(* IEC 61131-3 sources: 2026_Projet_YGO_ExcavatriceDragage/CODE_BACKUP/CODE_20260904_AvantWeekendBackup_v0.6.34/H_TREUILS_BENNE/_TYPES, 19 files *)

(* ---- E_WinchFinalInterlockReason.st ---- *)
(* =======================================================================
   🔒 E_WinchFinalInterlockReason — Raisons de blocage barrière finale
   ───────────────────────────────────────────────────────────────
   🎯 Rôle : Énumération des causes de neutralisation/interlock final treuil
   📄 Doc métier : DOC/AF/AF_Partie-10_Fonction_Winch_v2.1.md
   ======================================================================= *)
{attribute 'qualified_only'}
TYPE E_WinchFinalInterlockReason :
(
    NONE                        := 0,                                 // Aucun blocage actif
    BRAKE_COMMAND_NOT_CONFIRMED := 1,                                 // Absence confirmation ouverture frein > 500ms
    RESTART_INHIBITED           := 2,                                 // Inhibition redemarrage actif
    SENSE_DROP_TIMEOUT          := 3                                  // T_max §3bis depasse sans confirmation retombee (AC7)
);
END_TYPE

(* ---- E_WinchFinalInterlockState.st ---- *)
(* =======================================================================
   ⚙️ E_WinchFinalInterlockState — États machine barrière finale treuil
   ───────────────────────────────────────────────────────────────
   🎯 Rôle : Énumération des états opérationnels de l'interlock final
   📄 Doc métier : DOC/AF/AF_Partie-10_Fonction_Winch_v2.1.md
   ======================================================================= *)
{attribute 'qualified_only'}
TYPE E_WinchFinalInterlockState :
(
    DISABLED                        := 0,                             // Desactive / Hors service
    READY                           := 1,                             // Pret / Etat nominal
    WAIT_BRAKE_COMMAND_CONFIRMATION := 2,                             // Attente confirmation feedback frein
    WAIT_STEP_DELAY                 := 3,                             // Temporisation changement de palier
    WAIT_RESTART_DELAY              := 4,                             // Temporisation anti-court-cycle redemarrage
    FAULT                           := 5,                             // Etat de defaut
    WAIT_SENSE_DROP_CONFIRM         := 6                              // Maintien §3bis du contacteur de sens (AC6/AC7)
);
END_TYPE

(* ---- ST_fbBucketCmdArbitration_Context.st ---- *)
(* ═══════════════════════════════════════════════════════════════
   🧩 ST_fbBucketCmdArbitration_Context — Contexte de gating benne
   ───────────────────────────────────────────────────────────────
   🎯 Rôle : Encapsuler les faits de gating consommés par FB_BucketCmdArbitration
       pour le séquencement couplé benne (config, intention both, état benne).
       Le FB dérive les flags armés (WinchBothDiveBucketOpenArmed /
       WinchBothAscentBucketCloseArmed) et les commandes arbitrées.
   📤 Producteur : PRG_04_Treuils_Benne (câblage).
   📄 Doc : DOC/AF/AF_Partie-10_Fonction_Winch_v2.1.md
   🔌 État benne : 2 bits BOOL (BucketIsOpen/Closed) dérivés de _BucketState.
   ═══════════════════════════════════════════════════════════════ *)

TYPE ST_fbBucketCmdArbitration_Context :
STRUCT
    TglEnableCoupledBucketSequencing : BOOL;  // --> [CFG] Activation séquencement couplé benne (Commun.Cfg)
    MotionActive                     : BOOL;  // --> [CMD] Intention mouvement both active (WinchBothMotionActive)
    ReqAscent                        : BOOL;  // --> [CMD] Intention both montée
    ReqDescend                       : BOOL;  // --> [CMD] Intention both descente
    BucketIsOpen                     : BOOL;  // --> [STAT] Benne ouverte (BucketState.IsOpen)
    BucketIsClosed                   : BOOL;  // --> [STAT] Benne fermée (BucketState.IsClosed)
    CoupledPhaseLocked               : BOOL;  // --> [STAT] T248 : phase couplée verrouillée (Auth.CoupledBucketPhaseLocked) -> ne PAS (ré)armer dive-open/ascent-close : plus de correction benne ni de blocage sur l'état temps réel une fois le mouvement lancé
END_STRUCT
END_TYPE

(* ---- ST_fbBucketCmdArbitration_IHM.st ---- *)
(* ═══════════════════════════════════════════════════════════════
   🎛️ ST_fbBucketCmdArbitration_IHM — Entrées IHM de l'arbitrage benne
   ───────────────────────────────────────────────────────────────
   🎯 Rôle : Encapsuler les commandes IHM consommées par FB_BucketCmdArbitration
       (boutons ouverture/fermeture benne, nommage hardware propagé).
   📤 Producteur : PRG_04_Treuils_Benne (câblage GVL_IHM).
   📄 Doc : DOC/AF/AF_Partie-10_Fonction_Winch_v2.1.md
   🔌 Nommage : BtnOpen/BtnClose = nommage hardware propagé (convention projet).
   ═══════════════════════════════════════════════════════════════ *)

TYPE ST_fbBucketCmdArbitration_IHM :
STRUCT
    BtnOpen  : BOOL;  // --> [CMD] Bouton ouverture benne (M2TreuilBenne.Bucket.Cmd.BtnOpen)
    BtnClose : BOOL;  // --> [CMD] Bouton fermeture benne (M2TreuilBenne.Bucket.Cmd.BtnClose)
END_STRUCT
END_TYPE

(* ---- ST_fbWinch_Cfg.st ---- *)
(* =======================================================================
   🪝 ST_fbWinch_Cfg — Configuration statique d'un treuil
   ───────────────────────────────────────────────────────────────
   🎯 Rôle : Réglages persistants propres à l'instance treuil (statique)
   📄 Doc métier : DOC/AF/AF_Partie-10_Fonction_Winch_v2.1.md
   📤 Producteur : configuration persistante
   📥 Consommateur : FB_Winch (statique uniquement)
   🔒 Structs cibles + champs conservés pour garder le décodage %→palier
      et les deux cadences de rampe DANS FB_Winch (comportement
      bit-identique). Le champ StepRampDelay est déclaré mais non
      consommé (usage aval).
   ======================================================================= *)
TYPE ST_fbWinch_Cfg :
STRUCT
    // === TABLE DES PALIERS ===
    SpeedStepTable                  : ST_SpeedStepTable;   // Table de seuils des paliers de vitesse

    // === INTERLOCK CHANGEMENT DE SENS ===
    DirectionInterlockDelayAscent       : TIME := T#900ms;   // Delai interlock changement de sens montee
    DirectionInterlockDelayDescent     : TIME := T#400ms;   // Delai interlock changement de sens descente

    // === CADENCE DE RAMPE PALIER ===
    StepRampDelay                   : TIME := T#1000ms;  // [cible] Tempo de rampe palier (usage aval)
    StepRampDelayAscent             : TIME := T#1000ms;  // [08a] Cadence palier montee (D10, dedie)
    StepRampDelayDescent         : TIME := T#500ms;   // [08a] Cadence palier descending (D10, dedie)

    // === RETOMBÉE CONTACTEURS ===
    ContactorFeedbackTimeout        : TIME := T#500ms;   // Delai d'attente retombee des contacteurs

    // === RALENTISSEMENT BORDURE ===
    SlowdownDistanceTop_M           : REAL := 0.0;   // Distance avant limite haute pour ralentir (m) : 0 = arrêt au seuil
    SlowdownDistanceBottom_M        : REAL := 1.0;   // Distance avant limite basse pour ralentir (m)
    SlowdownMaxStep                 : INT := 1;      // Plafond palier dans zone de ralentissement (1..5)

    // === DÉCODAGE %→PALIER (conservé) ===
    SpeedStepHystMargin             : REAL := 2.0;   // [08a] Marge d'hysteresis palier (%)
END_STRUCT
END_TYPE

(* ---- ST_fbWinch_DriveRequest.st ---- *)
(* =======================================================================
   🪝 ST_fbWinch_Req — Requête d'axe treuil (producteur PRG_04)
   ───────────────────────────────────────────────────────────────
   🎯 Rôle : Demande de mouvement, palier et bornes de clamp d'un treuil
   📄 Doc métier : DOC/AF/AF_Partie-10_Fonction_Winch_v2.1.md
   📤 Producteur : PRG_04_Treuils_Benne (une par treuil M1/M2)
   📥 Consommateur : FB_Winch
   🔒 Structs cibles + champs conservés pour garder le décodage %→palier
      et le clamp DANS FB_Winch (comportement bit-identique).
      SpeedStepReq est consommé par FB_Winch (§5) ; MinStepUp est déclaré
      mais non consommé (usage aval).
   ======================================================================= *)
TYPE ST_fbWinch_Req :
STRUCT
    // === ORDRE DE MOUVEMENT ===
    RunRequest                      : BOOL;   // TRUE = mouvement demandé
    ReqAscent                       : BOOL;   // TRUE = demande montée
    ReqDescend                      : BOOL;   // TRUE = demande descente
    SpeedStepReq                    : INT;    // [cible] Palier demandé (1..5, 0 = arrêt) — consommé par FB_Winch

    // === BORNES DE CLAMP (agrégées PRG_04) ===
    MinStepUp                       : INT;    // [cible] Plancher palier montée (usage aval)
    MaxStepUp                       : INT := 5;    // Plafond palier montée (1..5)
    MinStepDown                     : INT := 0;    // Plancher palier descente (0 = aucun) -- plongee Kobold
    MaxStepDown                     : INT := 3;    // Plafond palier descente (1..5)

    // === LIMITES EFFECTIVES DU CYCLE ===
    TopLimitM                       : REAL := 8.5;   // Position limite haute active (m)
    BottomLimitM                    : REAL := -20.0; // Position limite basse active (m)

    // === DIAGNOSTIC (jamais lu par la logique FB_Winch) ===
    SyncCoupled                     : BOOL;   // [diag] Couplage synchro actif (garde de revue)

    // === CHAMPS CONSERVÉS (clamp interne FB_Winch) ===
    HomingApproachActive            : BOOL;   // [08a] Vitesse limitée au palier 1 (approche homing)
END_STRUCT
END_TYPE

(* ---- ST_fbWinch_Sensors.st ---- *)
(* =======================================================================
   🪝 ST_fbWinch_Sensors — Mesures et feedbacks d'un treuil
   ───────────────────────────────────────────────────────────────
   🎯 Rôle : Retours physiques et mesures propres à l'instance treuil
   📄 Doc métier : DOC/AF/AF_Partie-10_Fonction_Winch_v2.1.md
   📤 Producteur : PRG_04_Treuils_Benne / acquisition
   📥 Consommateur : FB_Winch
   🔒 Structs cibles + champs conservés pour garder le garde-fou vitesse
      DANS FB_Winch (comportement bit-identique). Les champs
      MeasuredSpeedMps / MeasuredSpeedValid sont déclarés mais non
      consommés (usage aval).
   ======================================================================= *)
TYPE ST_fbWinch_Sensors :
STRUCT
    // === POSITION ET RÉFÉRENCEMENT ===
    CablePosM                       : REAL;   // Position actuelle du cable (m)
    Homed                           : BOOL;   // Statut treuil reference
    HomingSuspect                   : BOOL;   // Incertitude / doute sur le referencement

    // === RETOURS CONTACTEURS ===
    ContactorsAllOff                : BOOL;   // TRUE = relais sens + C1..C4 tous retombés (ex-FwdRevSpeedFeedbackOff)

    // === MESURE VITESSE ===
    MeasuredSpeedMps                : REAL;   // [cible] Mesure vitesse réelle (m/s) — usage aval
    MeasuredSpeedValid              : BOOL;   // [cible] Mesure exploitable — usage aval
    MeasuredSpeedBand               : INT := 0;   // [08a] Bande vitesse réelle validée (garde-fou conservé dans FB_Winch)

    // === GARDE-FOU VITESSE (conservé) ===
    SpeedGuardEnable                : BOOL := TRUE;   // [08a] Activation garde-fou changement de palier
    SpeedGuardReady                 : BOOL := FALSE;  // [08a] Conditions de stabilité validées
END_STRUCT
END_TYPE

(* ---- ST_fbWinch_Symmetry_Cfg.st ---- *)
(* =======================================================================
   ⚖️ ST_fbWinch_Symmetry_Cfg — Configuration des seuils de symétrie M1/M2
   ───────────────────────────────────────────────────────────────
   🎯 Rôle : Seuils de tolérance pour le diagnostic passif de symétrie treuils
   📄 Doc métier : DOC/AF/AF_Partie-10_Fonction_Winch_v2.1.md
   ======================================================================= *)
TYPE ST_fbWinch_Symmetry_Cfg :
STRUCT
    DeltaStartDelay_Ms       : UDINT := 100;                          // Ecart max tolere au demarrage (ms)
    DeltaBrakeReleaseTime_Ms : UDINT := 100;                          // Ecart max temps desserrage frein (ms)
    DeltaBrakeApplyTime_Ms   : UDINT := 100;                          // Ecart max temps serrage frein (ms)
    DeltaStopDistance_Mm     : UDINT := 100;                          // Ecart max distance d'arret (mm)
    DeltaStopTime_Ms         : UDINT := 200;                          // Ecart max temps d'arret (ms)
    MinimumCommandTime_Ms    : UDINT := 1000;                         // Duree minimale de commande pour qualification (ms)
    MinimumSpeed_Mps         : REAL  := 0.05;                         // Vitesse minimale pour qualification (m/s)
END_STRUCT
END_TYPE

(* ---- ST_fbWinch_Symmetry_Data.st ---- *)
(* =======================================================================
   📊 ST_fbWinch_Symmetry_Data — Données mesurées de symétrie M1/M2
   ───────────────────────────────────────────────────────────────
   🎯 Rôle : Structure des résultats de mesures et d'écarts du diagnostic symétrie
   📄 Doc métier : DOC/AF/AF_Partie-10_Fonction_Winch_v2.1.md
   ======================================================================= *)
TYPE ST_fbWinch_Symmetry_Data :
STRUCT
    DeltaStartDelay_Ms       : UDINT;                                 // Ecart mesure au demarrage (ms)
    DeltaBrakeReleaseTime_Ms : UDINT;                                 // Ecart mesure temps desserrage frein (ms)
    DeltaBrakeApplyTime_Ms   : UDINT;                                 // Ecart mesure temps serrage frein (ms)
    DeltaStopDistance_Mm     : UDINT;                                 // Ecart mesure distance d'arret (mm)
    DeltaStopTime_Ms         : UDINT;                                 // Ecart mesure temps d'arret (ms)
    MaxSyncDeviation_M       : REAL;                                  // Ecart maximal de synchronisme enregistre (m)
END_STRUCT
END_TYPE

(* ---- ST_fbWinchCmdArbitration_Cfg.st ---- *)
(* ═══════════════════════════════════════════════════════════════
   ⚙️ ST_fbWinchCmdArbitration_Cfg — Config treuil (partagé M1/M2)
   ───────────────────────────────────────────────────────────────
   🎯 Rôle : Config statique de FB_WinchCmdArbitrationM1/M2.
       Structure UNIQUE partagée : M1 consomme BtnStepTgt (boutons/both),
       M2 consomme BtnStepTgt (boutons/both) + BucketOverrideStepTgt (chemin benne).
   📤 Producteur : PRG_04_Treuils_Benne (câblage).
   📄 Doc : DOC/AF/AF_Partie-10_Fonction_Winch_v2.1.md
   🔌 Remplace les paliers codés en dur (StepTgt := 5 / StepTgt := 1) par des constantes nommées.
   ═══════════════════════════════════════════════════════════════ *)

TYPE ST_fbWinchCmdArbitration_Cfg :
STRUCT
    BtnStepTgt : INT := 5;  // --> [CFG] Palier boutons/both (100 % → palier max)
    BucketOverrideStepTgt : INT := 1;  // --> [CFG] Palier override benne (vitesse lente)
END_STRUCT
END_TYPE

(* ---- ST_fbWinchCmdArbitration_Context.st ---- *)
(* ═══════════════════════════════════════════════════════════════
   🧩 ST_fbWinchCmdArbitration_Context — Contexte de gating treuil (partagé M1/M2)
   ───────────────────────────────────────────────────────────────
   🎯 Rôle : Encapsuler les faits de gating consommés par FB_WinchCommandArbitrationM1/M2
       (benne, synchro, blocage both). Structure UNIQUE partagée par les 2 axes,
       identifiée par l'instance : M1 ignore le chemin benne, M2 le consomme.
   📤 Producteur : PRG_04_Treuils_Benne (câblage).
   📄 Doc : DOC/AF/AF_Partie-10_Fonction_Winch_v2.1.md
   🔌 Action benne : 2 bits BOOL directionnels M2 issus de FB_Bucket.
   ═══════════════════════════════════════════════════════════════ *)

TYPE ST_fbWinchCmdArbitration_Context :
STRUCT
    BucketBusy                     : BOOL;  // --> [STAT] Action benne en cours (instBucket.Lifecycle.Busy)
    BucketM2RunRequest             : BOOL;  // --> [CMD] Commande M2 par la benne active
    BucketM2ReqAscent              : BOOL;  // --> [CMD] Demande montée M2 issue benne
    BucketM2ReqDescend             : BOOL;  // --> [CMD] Demande descente M2 issue benne
    WinchBothMotionBlockedByBucket : BOOL;  // --> [STAT] Mouvement both bloqué par benne (ex CoupledMotionBlockedByBucket)
    SyncBlocksAscent                   : BOOL;  // --> [STAT] Synchro bloque la montée (SyncMinorDeviationBlocksUp)
    SyncBlocksDescent                 : BOOL;  // --> [STAT] Synchro bloque la descente (SyncMinorDeviationBlocksDown)

    // === 🔗 ATOMICITÉ DE LA COMMANDE BOTH : permis agrégés consommés ===
    // PRG_04 calcule BothAscentPermit/BothDescendPermit = AND des 4 permits effectifs.
    // En commande both, la commande ne consomme QUE ces agrégats (jamais les permits
    // individuels directement) : les 2 treuils partent ensemble ou aucun (NC-100).
    M1AscentAllowed                 : BOOL;  // --> [SAFE] Fait EffectivePermitM1_Ascent
    M1DescendAllowed                : BOOL;  // --> [SAFE] Fait EffectivePermitM1_Descend
    M2AscentAllowed                 : BOOL;  // --> [SAFE] Fait EffectivePermitM2_Ascent
    M2DescendAllowed                : BOOL;  // --> [SAFE] Fait EffectivePermitM2_Descend
    BothBlock                       : BOOL;  // --> [STAT] Commande Both bloquée (aucun départ possible — diagnostic IHM)
END_STRUCT
END_TYPE

(* ---- ST_fbWinchCmdArbitration_IHM.st ---- *)
(* ═══════════════════════════════════════════════════════════════
   🎛️ ST_fbWinchCmdArbitration_IHM — Entrées IHM de l'arbitrage treuil
   ───────────────────────────────────────────────────────────────
   🎯 Rôle : Encapsuler les commandes IHM consommées par FB_WinchCommandArbitrationM1/M2
       (boutons par treuil, nommage hardware propagé).
       Le toggle joystick maître global (Modes.Cmd.TglJoystickMaster) est passé en
       paramètre séparé des FB (I4 — factorisation, source unique GVL_IHM.Modes.Cmd).
   📤 Producteur : PRG_04_Treuils_Benne (câblage GVL_IHM).
   📄 Doc : DOC/AF/AF_Partie-10_Fonction_Winch_v2.1.md
   🔌 Nommage : BtnAscentM1/BtnAscentM2 = nommage hardware propagé (convention projet).
   ═══════════════════════════════════════════════════════════════ *)

TYPE ST_fbWinchCmdArbitration_IHM :
STRUCT
    BtnAscentM1           : BOOL;  // --> [CMD] Bouton montée treuil M1 (nommage hardware)
    BtnDescentM1         : BOOL;  // --> [CMD] Bouton descente treuil M1
    BtnAscentM2           : BOOL;  // --> [CMD] Bouton montée treuil M2
    BtnDescentM2         : BOOL;  // --> [CMD] Bouton descente treuil M2
    BtnWinchBothAscent    : BOOL;  // --> [CMD] Bouton montée couplée both (Commun)
    BtnWinchBothDescent  : BOOL;  // --> [CMD] Bouton descente couplée both (Commun)
END_STRUCT
END_TYPE

(* ---- ST_fbWinchLoadEstimator_SpeedCfg.st ---- *)
(* =======================================================================
   ⚙️ ST_fbWinchLoadEstimator_SpeedCfg — Configuration des plages de vitesse linéaire
   ───────────────────────────────────────────────────────────────
   🎯 Rôle : Caractérisation des plages de vitesse mesurée par palier (m/s)
   📄 Doc métier : DOC/AF/AF_Partie-10_Fonction_Winch_v2.1.md
   ======================================================================= *)
TYPE ST_fbWinchLoadEstimator_SpeedCfg :
STRUCT
    MaxMeasuredSpeedMps    : REAL;                                    // Vitesse maximale mesuree de reference (m/s)
    SpeedBandMaxMps        : ARRAY[1..5] OF REAL;                    // Plafonds vitesse mesuree par palier (m/s)
    SpeedBandHysteresisMps : REAL;                                    // Hysteresis anti-battement classement vitesse (m/s)
END_STRUCT
END_TYPE

(* ---- ST_fbWinchLoadEstimator_Table.st ---- *)
(* =======================================================================
   📊 ST_fbWinchLoadEstimator_Table — Table empirique de charge estimée
   ───────────────────────────────────────────────────────────────
   🎯 Rôle : Matrice 5x5 d'estimation de charge (palier commandé x bande vitesse)
   📄 Doc métier : DOC/AF/AF_Partie-10_Fonction_Winch_v2.1.md
   ======================================================================= *)
TYPE ST_fbWinchLoadEstimator_Table :
STRUCT
    IsConfigured              : BOOL;                                 // Validation explicite de la table
    LoadPctByStepAndSpeedBand : ARRAY[1..5] OF ARRAY[1..5] OF REAL;  // Matrice [palier][bande_vitesse] charge (%)
END_STRUCT
END_TYPE

(* ---- ST_fbWinchSpeedLearning_Cell.st ---- *)
(* =======================================================================
   💾 ST_fbWinchSpeedLearning_Cell — Cellule de vitesse apprise
   ───────────────────────────────────────────────────────────────
   🎯 Rôle : Cellule unitaire de la table d'apprentissage vitesse par palier
   📄 Doc metier : DOC/AF/AF_Partie-10_Fonction_Winch_v2.1.md
   ======================================================================= *)
TYPE ST_fbWinchSpeedLearning_Cell :
STRUCT
    Valid       : BOOL;    // Cellule validee (vitesse apprise exploitable)
    SpeedMps    : REAL;    // Vitesse apprise (m/s)
    SampleCount : UDINT;   // Compteur d'echantillons collectes
END_STRUCT
END_TYPE

(* ---- ST_fbWinchSpeedLearning_Cfg.st ---- *)
(* =======================================================================
   ⚙️ ST_fbWinchSpeedLearning_Cfg — Enveloppes de plausibilite par palier
   ───────────────────────────────────────────────────────────────
   🎯 Rôle : Bornes min/max de vitesse apprise par palier + seuil d'echantillons
   📄 Doc metier : DOC/AF/AF_Partie-10_Fonction_Winch_v2.1.md
   ======================================================================= *)
TYPE ST_fbWinchSpeedLearning_Cfg :
STRUCT
    MinSpeedMps : ARRAY[1..5] OF REAL;   // Borne min vitesse apprise par palier (m/s)
    MaxSpeedMps : ARRAY[1..5] OF REAL;   // Borne max vitesse apprise par palier (m/s)
    MinSamples  : UDINT;                 // Nb min d'echantillons pour valider une cellule
END_STRUCT
END_TYPE

(* ---- ST_fbWinchSpeedLearning_Table.st ---- *)
(* =======================================================================
   💾 ST_fbWinchSpeedLearning_Table — Table RETAIN apprentissage vitesse
   ───────────────────────────────────────────────────────────────
   🎯 Rôle : Matrice {axe x sens x charge/vide x palier} de vitesses apprises
   📄 Doc metier : DOC/AF/AF_Partie-10_Fonction_Winch_v2.1.md
   ======================================================================= *)
TYPE ST_fbWinchSpeedLearning_Table :
STRUCT
    // [axe][sens][charge][palier]
    //   axe    : 1=M1, 2=M2
    //   sens   : 1=montee, 2=descente
    //   charge : 1=vide, 2=charge
    //   palier : 1..5
    Cell : ARRAY[1..2, 1..2, 1..2, 1..5] OF ST_fbWinchSpeedLearning_Cell;
END_STRUCT
END_TYPE

(* ---- ST_SpeedStepTable.st ---- *)
(* =======================================================================
   🪜 ST_SpeedStepTable — Table des paliers de vitesse contacteurs
   ───────────────────────────────────────────────────────────────
   🎯 Rôle : Structure de configuration des contacteurs et seuils par palier
   📄 Doc métier : DOC/AF/AF_Partie-10_Fonction_Winch_v2.1.md
   ======================================================================= *)
TYPE ST_SpeedStepTable :
STRUCT
    // === PALIER 1 (VITESSE MINIMALE) ===
    P1R1              : BOOL;                                         // Contacteur 1 pour Palier 1
    P1R2              : BOOL;                                         // Contacteur 2 pour Palier 1
    P1R3              : BOOL;                                         // Contacteur 3 pour Palier 1
    P1R4              : BOOL;                                         // Contacteur 4 pour Palier 1

    // === PALIER 2 ===
    P2R1              : BOOL;                                         // Contacteur 1 pour Palier 2
    P2R2              : BOOL;                                         // Contacteur 2 pour Palier 2
    P2R3              : BOOL;                                         // Contacteur 3 pour Palier 2
    P2R4              : BOOL;                                         // Contacteur 4 pour Palier 2

    // === PALIER 3 ===
    P3R1              : BOOL;                                         // Contacteur 1 pour Palier 3
    P3R2              : BOOL;                                         // Contacteur 2 pour Palier 3
    P3R3              : BOOL;                                         // Contacteur 3 pour Palier 3
    P3R4              : BOOL;                                         // Contacteur 4 pour Palier 3

    // === PALIER 4 ===
    P4R1              : BOOL;                                         // Contacteur 1 pour Palier 4
    P4R2              : BOOL;                                         // Contacteur 2 pour Palier 4
    P4R3              : BOOL;                                         // Contacteur 3 pour Palier 4
    P4R4              : BOOL;                                         // Contacteur 4 pour Palier 4

    // === PALIER 5 (VITESSE MAXIMALE) ===
    P5R1              : BOOL;                                         // Contacteur 1 pour Palier 5
    P5R2              : BOOL;                                         // Contacteur 2 pour Palier 5
    P5R3              : BOOL;                                         // Contacteur 3 pour Palier 5
    P5R4              : BOOL;                                         // Contacteur 4 pour Palier 5

    // === SEUILS DE TRANSITION (%) ===
    StepThreshold_Pct : ARRAY[1..5] OF REAL;                          // Seuils de changement de palier (0..100%)
END_STRUCT
END_TYPE

(* ---- ST_SyncContactorDiag.st ---- *)
(* =======================================================================
   🔀 ST_SyncContactorDiag — Diagnostic discordance contacteurs M1/M2
   ───────────────────────────────────────────────────────────────
   🎯 Rôle : dire EN CLAIR quel contacteur diverge entre M1 et M2 et à quel
      niveau on est (aucun / mismatch confirmé / escalade). Consommé par le
      bandeau IHM et le troubleshooting pour répondre « pourquoi ça bloque ».
   🔒 Bits nommés (pas de masque hexa, AF03 §4). Plusieurs bits peuvent être
      TRUE simultanément (toutes les divergences détectées).
   📄 Doc : DOC/AF/AF_Partie-10_Fonction_Winch_v2.1.md
   ======================================================================= *)
TYPE ST_SyncContactorDiag :
STRUCT
    RelayFwdMismatch : BOOL; // TRUE = relais montée M1 <> M2
    RelayRevMismatch : BOOL; // TRUE = relais descente M1 <> M2
    Step1Mismatch    : BOOL; // TRUE = contacteur palier 1 M1 <> M2
    Step2Mismatch    : BOOL; // TRUE = contacteur palier 2 M1 <> M2
    Step3Mismatch    : BOOL; // TRUE = contacteur palier 3 M1 <> M2
    Step4Mismatch    : BOOL; // TRUE = contacteur palier 4 M1 <> M2
    MismatchLevel    : INT;  // 0 = aucun · 1 = discordance confirmée (SafeStop) · 2 = escalade (PowerCutOff)
END_STRUCT
END_TYPE
